// TIA Portal project "SludeProcess_Near_Final" (V16)

(* hardware
DEVICE "S71500/ET200MP station_1"  S7-1500 station
   slot 0: "Rail_0"  Rack  6ES7 590-1***0-0AA0
   slot 1: "PLC_1"  CPU 1511-1 PN  6ES7 511-1AK01-0AB0  V2.8
      slot 3: "CPU display_1"  6ES7591-1AA00-0AA0
      slot 32768: "PROFINET interface_1"  X1
         slot 32769: "Port_1"  X1 P1
         slot 32770: "Port_2"  X1 P2
      slot 34817: "Virtual CP interface port_1"  Virtual CP interface port  Virtual CP interface port
   slot 2: "DI 16x24VDC BA_1"  DI 16x24VDC BA  6ES7 521-1BH10-0AA0  V1.1
   slot 3: "DQ 16x24VDC/0.5A BA_1"  DQ 16x24VDC/0.5A BA  6ES7 522-1BH10-0AA0  V1.1
   slot 4: "AI 8xU/I/RTD/TC ST_1"  AI 8xU/I/RTD/TC ST  6ES7 531-7KF00-0AB0  V2.2
   slot 5: "AQ 2xU/I ST_1"  AQ 2xU/I ST  6ES7 532-5NB00-0AB0  V1.0
   slot 6: "DI 16x24VDC BA_2"  DI 16x24VDC BA  6ES7 521-1BH10-0AA0  V1.1
DEVICE "HMI_1"  KTP700 Basic PN
   slot 0: "HMI_1"  KTP700 Basic PN  6AV2 123-2GB03-0AX0  16.0.0.0
   slot 1: "HMI_RT_1"  KTP700 Basic PN  6AV2 123-2GB03-0AX0  16.0.0.0
   slot 5: "HMI_1.IE_CP_1"  PROFINET Interface  16.0.0.0
      slot 1: "PROFINET Interface_1"  PROFINET Interface
         slot 1: "Port_1"  Port
*)

// ===== PLC "PLC_1"  CPU 1511-1 PN =====

VAR_GLOBAL   // PLC tag table "Default tag table"
   "M001start" AT %M2.0 : Bool;
   "M001stop" AT %M12.1 : Bool;
   "FT-516_l/s" AT %MD12 : Real;
   "FT-516_status" AT %MW16 : Word;
   "FIC-516_setpoint" AT %MD18 : Real;
   "FIC-516_reset" AT %M2.1 : Bool;
   "M003_status" AT %MW20 : Word;
   "Test_open_valves" AT %M2.2 : Bool;
   "Test_M003_start" AT %M2.3 : Bool;
   "LT-515_liters" AT %MD22 : Real;
   "LT-515_status" AT %MW24 : Word;
   "M002_startbutton" AT %M2.4 : Bool;
   "M002_stopbutton" AT %M2.5 : Bool;
   "M002start" AT %M2.6 : Bool;
   "M002stop" AT %M2.7 : Bool;
   "WT-512_kg" AT %MD26 : Real;
   "TT-517_C" AT %MD28 : Real;
   "TT-518_C" AT %MD32 : Real;
   "WT-512_status" AT %MW36 : Word;
   "TT-517_status" AT %MW38 : Word;
   "TT-518_status" AT %MW40 : Word;
   "StartButton" AT %M3.0 : Bool;
   "StopButton" AT %M3.1 : Bool;
   "mixing" AT %M3.2 : Bool;
   "LSA513_HighLevel" AT %M3.3 : Bool;
   "HS519_FlowSwitch" AT %M3.4 : Bool;
   "HS514_MixReady" AT %M3.5 : Bool;
   "HS510_Valve" AT %M3.6 : Bool;
   "HS511_Valve" AT %M3.7 : Bool;
   "HS514_Valve" AT %M4.0 : Bool;
   "HS519_Valve" AT %M4.1 : Bool;
   "HS521_Alarm" AT %M4.2 : Bool;
   "M001_pMotor" AT %M4.3 : Bool;
   "M002_mix" AT %M4.4 : Bool;
   "M003_transferPump" AT %M4.5 : Bool;
   "FrequencyCommand" AT %MD42 : Real;
   "CurrentStep" AT %MW46 : Int;
   "Alarm" AT %M4.6 : Bool;
   "Step" AT %MW48 : Int;
   "NextStep" AT %MW50 : Int;
   "ResetButton" AT %M5.0 : Bool;
   "EmergencyButton" AT %M5.1 : Bool;
   "prevStart" AT %M5.2 : Bool;
   "prevStop" AT %M5.3 : Bool;
END_VAR

VAR_GLOBAL   // PLC tag table "SIMIT interface"
   "ZSO-510" AT %I0.0 : Bool;
   "ZSC-510" AT %I0.1 : Bool;
   "ZSO-511" AT %I0.2 : Bool;
   "ZSC-511" AT %I0.3 : Bool;
   "ZSO-514" AT %I0.4 : Bool;
   "ZSC-514" AT %I0.5 : Bool;
   "ZSO-519" AT %I0.6 : Bool;
   "ZSC-519" AT %I0.7 : Bool;
   "ZSO-521" AT %I1.0 : Bool;
   "ZSC-521" AT %I1.1 : Bool;
   "M001.R" AT %I1.2 : Bool;
   "M002.R" AT %I1.3 : Bool;
   "LS-513" AT %I1.4 : Bool;
   "GSV-510" AT %Q0.0 : Bool;
   "GSV-511" AT %Q0.1 : Bool;
   "GSV-514" AT %Q0.2 : Bool;
   "GSV-519" AT %Q0.3 : Bool;
   "GSV-521" AT %Q0.4 : Bool;
   "M001.ST" AT %Q0.5 : Bool;
   "M002.ST" AT %Q0.6 : Bool;
   "WT-512" AT %IW2 : Int;
   "LT-515" AT %IW4 : Int;
   "FT-516" AT %IW6 : Int;
   "TT-517" AT %IW8 : Int;
   "TT-518" AT %IW10 : Int;
   "M003.SP" AT %QW2 : Int;
   "M001.F" AT %I1.5 : Bool;
   "M002.F" AT %I1.6 : Bool;
   "M003.R" AT %I1.7 : Bool;
   "M003.F" AT %I18.0 : Bool;
   "M003.ST" AT %Q0.7 : Bool;
   "M001.TK" AT %I18.1 : Bool;
   "M002.TK" AT %I18.2 : Bool;
   "M003.TK" AT %I18.3 : Bool;
END_VAR

DATA_BLOCK "fb_ProcessSequence1_DB"   // DB2
{ S7_Optimized_Access := 'TRUE' }
VERSION : 0.1
// stored: InstanceOfName fb_ProcessSequence1
"fb_ProcessSequence1"
BEGIN
END_DATA_BLOCK

DATA_BLOCK "FIC516_DB"   // DB3
{ S7_Optimized_Access := 'TRUE' }
VERSION : 0.1
// stored: InstanceOfName FIC516
"FIC516"
BEGIN
END_DATA_BLOCK

DATA_BLOCK "AI_handeling_DB"   // DB14
{ S7_Optimized_Access := 'TRUE' }
VERSION : 0.1
// stored: InstanceOfName AI_handeling
"AI_handeling"
BEGIN
END_DATA_BLOCK

// folder: System blocks/Program resources

DATA_BLOCK "tMix"   // DB4
{ S7_Optimized_Access := 'TRUE' }
AUTHOR : Simatic
FAMILY : IEC
NAME : IEC_TMR
VERSION : 1.0
// stored: InstanceOfName IEC_TIMER
"IEC_TIMER"
BEGIN
END_DATA_BLOCK

// folder: (top level)

FUNCTION_BLOCK "FIC516"   // FB1, FBD
{ S7_Optimized_Access := 'TRUE' }
VERSION : 0.1
BEGIN

REGION Network 1
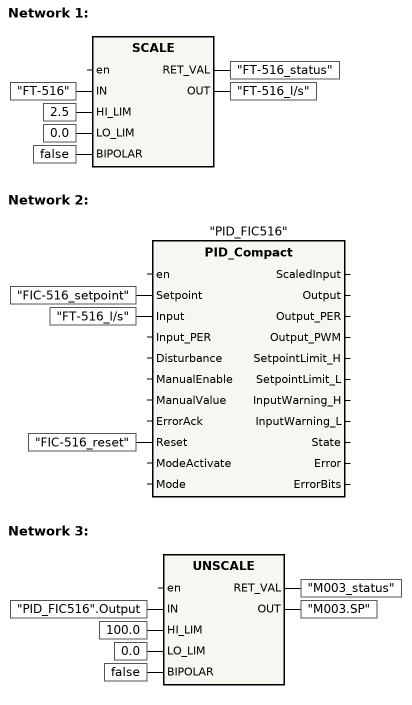
   "FT-516_status" := SCALE(IN := "FT-516", HI_LIM := 2.5, LO_LIM := 0.0, BIPOLAR := false, OUT => "FT-516_l/s");
END_REGION

REGION Network 2
   "PID_FIC516"(Setpoint := "FIC-516_setpoint", Input := "FT-516_l/s", Reset := "FIC-516_reset");   // PID_Compact
END_REGION

REGION Network 3
   "M003_status" := UNSCALE(IN := "PID_FIC516".Output,
                           HI_LIM := 100.0,
                           LO_LIM := 0.0,
                           BIPOLAR := false,
                           OUT => "M003.SP");
END_REGION
END_FUNCTION_BLOCK

FUNCTION_BLOCK "AI_handeling"   // FB4, FBD
{ S7_Optimized_Access := 'TRUE' }
VERSION : 0.1
BEGIN

REGION Network 1
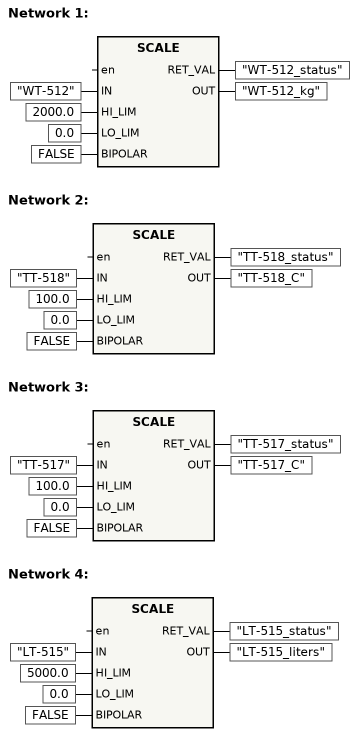
   "WT-512_status" := SCALE(IN := "WT-512",
                           HI_LIM := 2000.0,
                           LO_LIM := 0.0,
                           BIPOLAR := FALSE,
                           OUT => "WT-512_kg");
END_REGION

REGION Network 2
   "TT-518_status" := SCALE(IN := "TT-518", HI_LIM := 100.0, LO_LIM := 0.0, BIPOLAR := FALSE, OUT => "TT-518_C");
END_REGION

REGION Network 3
   "TT-517_status" := SCALE(IN := "TT-517", HI_LIM := 100.0, LO_LIM := 0.0, BIPOLAR := FALSE, OUT => "TT-517_C");
END_REGION

REGION Network 4
   "LT-515_status" := SCALE(IN := "LT-515",
                           HI_LIM := 5000.0,
                           LO_LIM := 0.0,
                           BIPOLAR := FALSE,
                           OUT => "LT-515_liters");
END_REGION
END_FUNCTION_BLOCK

FUNCTION_BLOCK "fb_ProcessSequence1"   // FB5, SCL
{ S7_Optimized_Access := 'TRUE' }
VERSION : 0.1
   VAR_INPUT
      StartButton : Bool := false;
      StopButton : Bool;
      RestartButton : Bool;
      ResetButton : Bool;
      EmergencyButton : Bool;
      "WT-512_kg" : Real;
      LT_515_liters : Real;
      FIC_516_setpoint : Real;
      TT_517_C : Real;
      TT_518_C : Real;
      LSA513_HighLevel : Bool;
      HS519_FlowSwitch : Bool;
      HS514_MixReady : Real;
      M001_SafetySwitch : Bool;
      M002_SafetySwitch : Bool;
      M003_SafetySwitch : Bool;
      Mode_Manual : Bool;
   END_VAR
   VAR_OUTPUT
      HS514_Valve : Bool;
      HS510_Valve : Bool;
      HS511_Valve : Bool;
      HS519_Valve : Bool;
      HS521_Valve : Bool;
      M001_pMotor : Bool;
      M002_mix : Bool;
      M003_TransferPump : Bool;
      FrequencyCommand : Real;
   END_VAR
   VAR
      Filling : Bool;
      WeightSetpoint : Real := 800.0;
      prevStart : Bool;
      AlarmActive : Bool;
      DosingNaOH : Bool;
      FeedingPowder : Bool;
      prevStop : Bool;
      Mixing : Bool;
      Transferring : Bool;
      StepMem : Bool;
      tMixTimer : Time;
      tFlowTimer : Time;
      "Step" : Int;
      Mode_Auto : Bool := true;
      HS519_manualValve : Bool;
      CircActive : Bool := false;
      MAN_HS510 : Bool;
      MAN_HS511 : Bool;
      MAN_HS514 : Bool;
      MAN_M001 : Bool;
      MAN_M002 : Bool;
      MAN_M003 : Bool;
      paused : Bool;
      M002_Fault_1 : Bool;
      restartLatch : Bool;
      TT_517_alarm : Bool;
      TT_518_alarm : Bool;
      LSA_513 : Bool := true;
      M001_Fault : Bool;
      M002_Fault : Bool;
      M003_Fault : Bool;
      CurrentStep : Int;
      Alarm : Bool;
      AlarmCause : String;
      M001_Safety : Bool;
      M002_Safety : Bool;
      M003_Safety : Bool;
      cMixTime : Time := T#20s;
      cOpenValveTime : Time := T#1000ms;
      cFlowCtrlTime : Time := T#50ms;
      running : Bool;
   END_VAR
   VAR CONSTANT
      cWeightWater : Real := 800.0;
      cWeightNaOH : Real := 1500.0;
      cWeightPowder : Real := 1000.0;
      cMaxWeight : Real := 2500.0;
      cFlowMin : Real := 0.5;
      cFlowMax : Real := 2.5;
      cTempEmergency : Real := 150.0;
      cTransferTrip : Real := 40.0;
      cFrequencyStep : Real := 1.0;
      cFrequenceMax : Real := 100.0;
      cFrequencyMin : Real;
   END_VAR
BEGIN
   // ---------- Immediate Emergency & Interlocks ----------
   IF #EmergencyButton OR (#TT_517_C >= #cTempEmergency) OR (#"WT-512_kg" >= #cMaxWeight) THEN
       #Alarm := TRUE;
       #AlarmCause := 'Emergency Stop or Max Temp/Weight Exceeded';
       #HS510_Valve := FALSE;
       #HS511_Valve := FALSE;
       #HS514_Valve := FALSE;
       #HS519_Valve := FALSE;
       #HS521_Valve := FALSE;
       #M001_pMotor := FALSE;
       #M002_mix := FALSE;
       #M003_TransferPump := FALSE;
       #FrequencyCommand := 0.0;
       #Step := 99;
       #paused := FALSE;
       RETURN;
   END_IF;

   // ---------- Default Outputs & HMI Indicators Initialization ----------
   // Hardware Outputs
   #HS510_Valve := FALSE;
   #HS511_Valve := FALSE;
   #HS514_Valve := FALSE;
   #HS519_Valve := FALSE;
   #HS521_Valve := FALSE;
   #M001_pMotor := FALSE;
   #M002_mix := FALSE;
   #M003_TransferPump := FALSE;
   #FrequencyCommand := 0.0;

   // HMI Status Indicators (Reset every scan, forced ON during active steps)
   #Filling := FALSE;
   #FeedingPowder := FALSE;
   #DosingNaOH := FALSE;
   #Mixing := FALSE;
   #Transferring := FALSE;
   #running := FALSE;

   // Automatic detection of motor faults & Alarms
   IF #TT_517_C >= #cTempEmergency THEN
       #TT_517_alarm := TRUE;
   END_IF;
   IF #TT_517_alarm THEN
       #M002_Fault := TRUE;
       #M002_Safety := FALSE;
       #Alarm := TRUE;
       #AlarmCause := 'TI-517 overtemp -> M002 fault';
   END_IF;

   IF #TT_518_C >= #cTempEmergency THEN
       #TT_518_alarm := TRUE;
   END_IF;
   IF #TT_518_alarm THEN
       #M003_Fault := TRUE;
       #M003_Safety := FALSE;
       #Alarm := TRUE;
       #AlarmCause := 'TI-518 overtemp -> M003 fault';
   END_IF;

   // LSA 513 Powder Hopper Low Level Warning
   IF NOT #LSA513_HighLevel AND (#AlarmCause = '') THEN
       #AlarmCause := 'LSA_513 Powder Hopper Low Level Warning';
   END_IF;

   // Reset alarm 
   IF #ResetButton THEN
       #Alarm := FALSE;
       #M001_Fault := FALSE;
       #M002_Fault := FALSE;
       #M003_Fault := FALSE;
       #TT_517_alarm := FALSE;
       #TT_518_alarm := FALSE;
       #AlarmCause := '';
   END_IF;

   // Restart (Only functions AFTER alarms are cleared)
   IF #RestartButton AND NOT #EmergencyButton AND NOT #Alarm THEN
       IF #M001_Safety AND #M002_Safety AND #M003_Safety AND NOT #M001_Fault AND NOT #M002_Fault AND NOT #M003_Fault THEN
           #Step := 0;
           #FrequencyCommand := 0.0;
           #paused := FALSE;
       END_IF;
   END_IF;

   // Hardware Safety Switch Mapping (TRUE = Healthy Motor)
   #M001_Safety := #M001_SafetySwitch;
   #M002_Safety := #M002_SafetySwitch;
   #M003_Safety := #M003_SafetySwitch;

   // Delivery Request mapping
   IF #HS519_FlowSwitch THEN
       #HS519_manualValve := TRUE;
   ELSE
       #HS519_manualValve := FALSE;
   END_IF;

   // ---------- Manual mode ----------
   IF #Mode_Manual THEN
       #running := TRUE;
       #Mode_Auto := FALSE;

       IF #MAN_HS510 AND #M001_Safety AND #M002_Safety THEN
           #HS510_Valve := TRUE;
           #Filling := TRUE;
       END_IF;
       IF #MAN_HS511 AND #M002_Safety THEN
           #HS511_Valve := TRUE;
           #DosingNaOH := TRUE;
       END_IF;
       IF #MAN_HS514 THEN
           #HS514_Valve := TRUE;
           #Transferring := TRUE;
       END_IF;

       IF #MAN_M001 AND NOT #M001_Fault AND #M001_Safety THEN
           #M001_pMotor := TRUE;
           #FeedingPowder := TRUE;
       END_IF;

       IF #MAN_M002 AND NOT #M002_Fault AND #M002_Safety THEN
           #M002_mix := TRUE;
           #Mixing := TRUE;
       END_IF;

       IF #MAN_M003 AND NOT #M003_Fault AND #M003_Safety THEN
           #M003_TransferPump := TRUE;
       END_IF;

       GOTO Global_Interlocks;
   END_IF;


   // ---------- Auto Sequence Controls ----------
   IF #StopButton AND (NOT #prevStop) THEN
       #paused := NOT #paused; // rising edge toggle
   END_IF;
   IF #StartButton THEN
       #paused := FALSE;
   END_IF;
   #prevStop := #StopButton;

   IF #paused THEN
       #AlarmCause := 'Process PAUSED';
       GOTO Global_Interlocks;
   ELSE
       IF #AlarmCause = 'Process PAUSED' THEN
           #AlarmCause := '';
       END_IF;
   END_IF;


   // ==============================================================================
   // INDEPENDENT STORAGE TANK BACKGROUND CIRCULATION (Runs constantly in Auto Mode)
   // ==============================================================================
   IF #Mode_Auto AND (#Step <> 99) THEN
       IF #LT_515_liters > 500.0 THEN
           IF #M003_Safety AND NOT #M003_Fault THEN
               #M003_TransferPump := TRUE;
               #running := TRUE;

               IF #HS519_manualValve THEN
                   // Delivery Mode Active
                   #HS519_Valve := TRUE;
                   #HS521_Valve := FALSE;
                   #CircActive := FALSE;

                   // Flow Control logic
                   IF #FIC_516_setpoint > #cFlowMin AND #FIC_516_setpoint < #cFlowMax THEN
                       IF #FrequencyCommand < #FIC_516_setpoint THEN
                           #FrequencyCommand := MIN(IN1 := #FrequencyCommand + #cFrequencyStep, IN2 := #cFrequenceMax);
                       ELSIF #FrequencyCommand > #FIC_516_setpoint THEN
                           #FrequencyCommand := MAX(IN1 := #FrequencyCommand - #cFrequencyStep, IN2 := #cFrequencyMin);
                       END_IF;
                   END_IF;
               ELSE
                   // Default Recirculation Mode Active
                   #HS519_Valve := FALSE;
                   #HS521_Valve := TRUE;
                   #CircActive := TRUE;
               END_IF;
           ELSE
               #M003_TransferPump := FALSE;
               #CircActive := FALSE;
               #Alarm := TRUE;
               #AlarmCause := 'M003 unsafe for delivery/recirculation';
               #Step := 99;
           END_IF;
       END_IF;
   END_IF;
   // ==============================================================================


   // ---------- State Machine (Mix Tank Batching Sequence) ----------
   CASE #Step OF

       0: // Standby
           #Mode_Auto := TRUE;
           IF #StartButton THEN
               #Step := 2;
           END_IF;

       2: // Start Check
           #Mode_Auto := TRUE;
           IF #Mode_Auto THEN
               #Step := 3;
               "tMix".TON(IN := FALSE,
                          PT := #cMixTime); // Hard reset the timer so it is fresh for the new batch
           ELSE
               IF #StartButton THEN
                   #running := TRUE;
               END_IF;
           END_IF;

       3: // Water Dosing (HS 510)
           IF #M001_Safety AND NOT #M002_Fault THEN
               #HS510_Valve := TRUE;
               #running := TRUE;
               #Filling := TRUE;
           ELSE
               #Alarm := TRUE;
               #AlarmCause := 'Equipment unsafe for water fill';
               #Step := 99;
           END_IF;

           IF #"WT-512_kg" >= #cWeightWater THEN
               #Step := 4;
           END_IF;

       4: // Powder Dosing & Mixing (M001 & M002)
           IF #M001_Safety AND #M002_Safety AND NOT #M001_Fault AND NOT #M002_Fault THEN
               #M001_pMotor := TRUE;
               #M002_mix := TRUE;
               #FeedingPowder := TRUE;
               #Mixing := TRUE;
               #running := TRUE;
           ELSE
               #Alarm := TRUE;
               #AlarmCause := 'M001/M002 safety fault prevented powder feed';
               #Step := 99;
           END_IF;

           IF #"WT-512_kg" >= #cWeightPowder THEN
               #Step := 5;
           END_IF;

       5: // Sodium Hydroxide Dosing (HS 511 & M002)
           IF #M002_Safety AND NOT #M002_Fault THEN
               #HS511_Valve := TRUE;
               #M002_mix := TRUE;
               #DosingNaOH := TRUE;
               #Mixing := TRUE;
               #running := TRUE;
           ELSE
               #Alarm := TRUE;
               #AlarmCause := 'M002 unsafe during NaOH dosing';
               #Step := 99;
           END_IF;

           IF #"WT-512_kg" >= #cWeightNaOH THEN
               #Step := 6;
           END_IF;

       6: // Final Mixing Time (Waits for proper mix before transfer)
           IF #M002_Safety AND NOT #M002_Fault THEN
               #M002_mix := TRUE;
               #Mixing := TRUE;
               #running := TRUE;

               // Run the TON Timer
               "tMix".TON(IN := TRUE,
                          PT := #cMixTime,
                          ET => #tMixTimer);
           ELSE
               #Alarm := TRUE;
               #AlarmCause := 'M002 unsafe for final mixing';
               #Step := 99;
           END_IF;

           // Once the timer hits the PT value (e.g., 5s), Q goes TRUE
           IF "tMix".Q THEN
               "tMix".TON(IN := FALSE,
                          PT := #cMixTime); // Reset the timer before moving on
               #Step := 7;
           END_IF;

       7: // Transfer to Storage Tank (HS 514)
           IF #LT_515_liters < 4950.0 THEN
               #HS514_Valve := TRUE;
               #running := TRUE;
               #Transferring := TRUE;
           END_IF;

           // Sequence finishes when Mix Tank is empty. Goes straight back to Standby!
           IF (#"WT-512_kg" <= 10.0) OR (#LT_515_liters >= 4950.0) THEN
               #Step := 0;
           END_IF;

       99: // Fault State
           #running := FALSE;
           #CircActive := FALSE;

           // 1. Operator MUST press Reset first to clear the alarm
           IF #ResetButton THEN
               IF #M001_SafetySwitch AND #M002_SafetySwitch AND #M003_SafetySwitch AND NOT #M001_Fault AND NOT #M002_Fault AND NOT #M003_Fault THEN
                   #Alarm := FALSE; // Fault cleared successfully
                   #AlarmCause := '';
               ELSE
                   #Alarm := TRUE;
                   #AlarmCause := 'Cannot clear emergency - check faults/safety';
               END_IF;
           END_IF;

           // 2. ONLY after Reset clears the alarm, wait for Start or Restart command
           IF NOT #Alarm THEN
               IF #StartButton THEN
                   #Step := 2; // Press START to resume the batch from where it failed
               ELSIF #RestartButton THEN
                   #Step := 0; // Press RESTART to abort batch and return to Standby
               END_IF;
           END_IF;

       ELSE
           #Step := 0;
   END_CASE;

   // ---------- Global Interlocks (Applies to both Auto & Manual) ----------
   Global_Interlocks:

   // 1. Storage Tank Overflow Protection
   IF #LT_515_liters >= 4950.0 THEN
       #HS514_Valve := FALSE;
   END_IF;

   // 2. Storage Tank Low Level Pump Protection
   IF #LT_515_liters <= 500.0 THEN
       #M003_TransferPump := FALSE;
       #HS521_Valve := FALSE;
       #HS519_Valve := FALSE;
   END_IF;

   // 3. Flow Diverter Interlock: Cannot be open at the same time
   IF #HS519_Valve AND #HS521_Valve THEN
       #HS521_Valve := FALSE;
   END_IF;

   #CurrentStep := #Step;
END_FUNCTION_BLOCK

ORGANIZATION_BLOCK "Main"   // OB1, FBD, ProgramCycle
TITLE = "Main Program Sweep (Cycle)"
{ S7_Optimized_Access := 'TRUE' }
VERSION : 0.1
   VAR_INPUT
      Initial_Call : Bool;   // Initial call of this OB
      Remanence : Bool;   // =True, if remanent data are available
   END_VAR
BEGIN

REGION Network 1
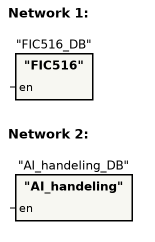
   "FIC516_DB"();   // "FIC516"
END_REGION

REGION Network 2
   "AI_handeling_DB"();   // "AI_handeling"
END_REGION

REGION Network 3
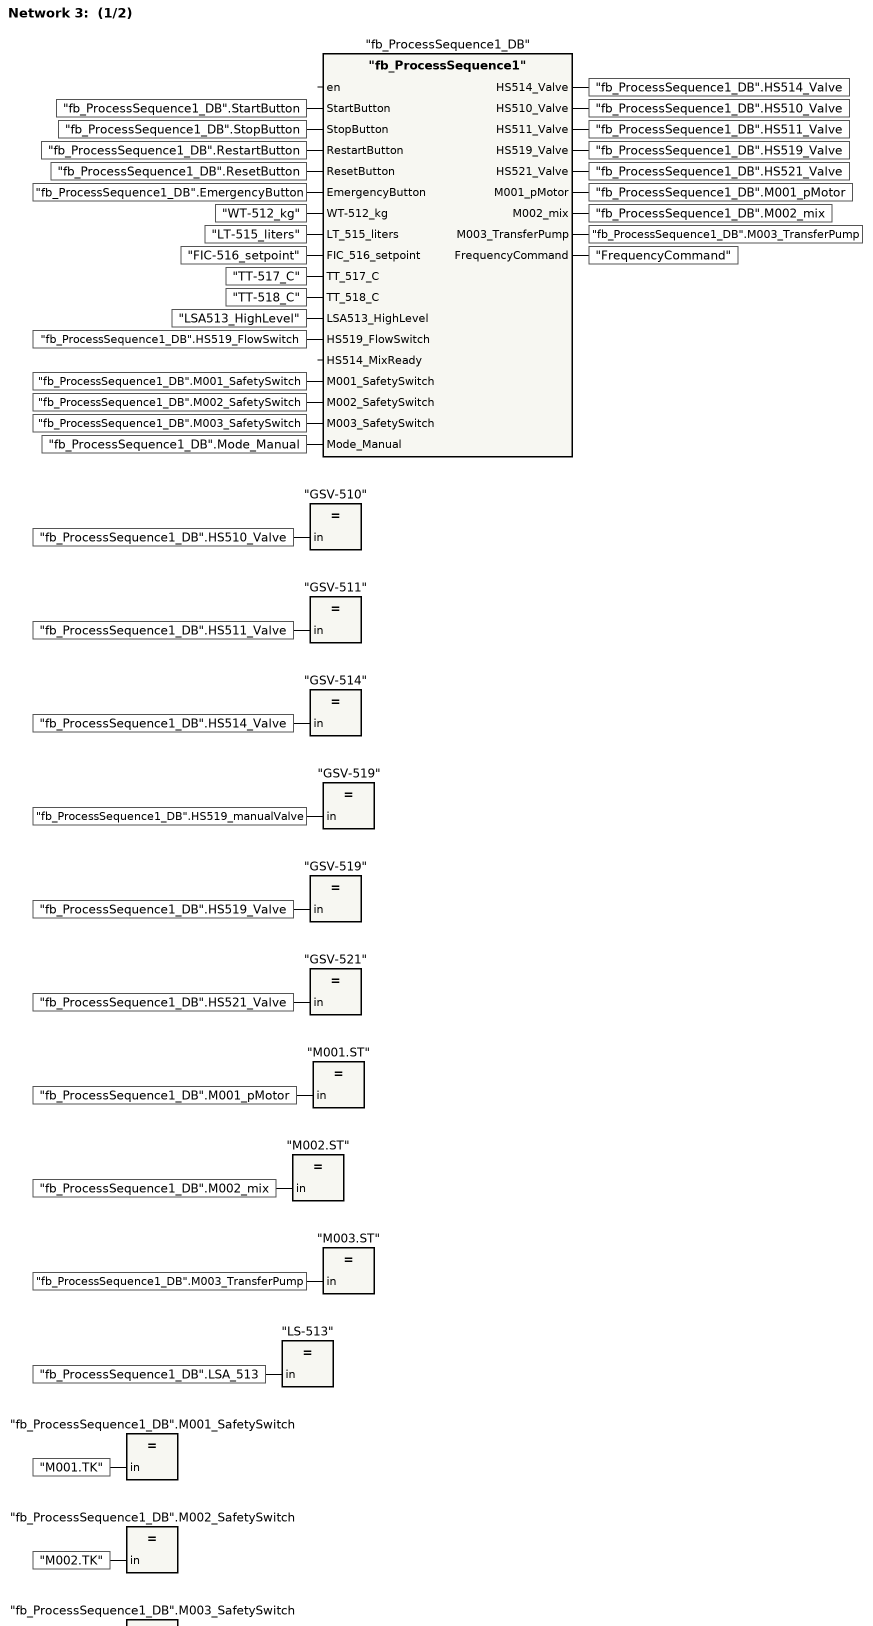
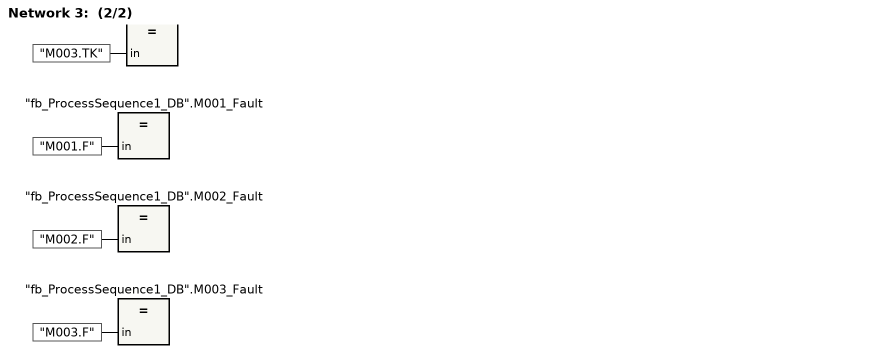
   "fb_ProcessSequence1_DB"(StartButton := "fb_ProcessSequence1_DB".StartButton,   // "fb_ProcessSequence1"
                           StopButton := "fb_ProcessSequence1_DB".StopButton,
                           RestartButton := "fb_ProcessSequence1_DB".RestartButton,
                           ResetButton := "fb_ProcessSequence1_DB".ResetButton,
                           EmergencyButton := "fb_ProcessSequence1_DB".EmergencyButton,
                           "WT-512_kg" := "WT-512_kg",
                           LT_515_liters := "LT-515_liters",
                           FIC_516_setpoint := "FIC-516_setpoint",
                           TT_517_C := "TT-517_C",
                           TT_518_C := "TT-518_C",
                           LSA513_HighLevel := "LSA513_HighLevel",
                           HS519_FlowSwitch := "fb_ProcessSequence1_DB".HS519_FlowSwitch,
                           M001_SafetySwitch := "fb_ProcessSequence1_DB".M001_SafetySwitch,
                           M002_SafetySwitch := "fb_ProcessSequence1_DB".M002_SafetySwitch,
                           M003_SafetySwitch := "fb_ProcessSequence1_DB".M003_SafetySwitch,
                           Mode_Manual := "fb_ProcessSequence1_DB".Mode_Manual,
                           HS514_Valve => "fb_ProcessSequence1_DB".HS514_Valve,
                           HS510_Valve => "fb_ProcessSequence1_DB".HS510_Valve,
                           HS511_Valve => "fb_ProcessSequence1_DB".HS511_Valve,
                           HS519_Valve => "fb_ProcessSequence1_DB".HS519_Valve,
                           HS521_Valve => "fb_ProcessSequence1_DB".HS521_Valve,
                           M001_pMotor => "fb_ProcessSequence1_DB".M001_pMotor,
                           M002_mix => "fb_ProcessSequence1_DB".M002_mix,
                           M003_TransferPump => "fb_ProcessSequence1_DB".M003_TransferPump,
                           FrequencyCommand => "FrequencyCommand");
   "GSV-510" := "fb_ProcessSequence1_DB".HS510_Valve;
   "GSV-511" := "fb_ProcessSequence1_DB".HS511_Valve;
   "GSV-514" := "fb_ProcessSequence1_DB".HS514_Valve;
   "GSV-519" := "fb_ProcessSequence1_DB".HS519_manualValve;
   "GSV-519" := "fb_ProcessSequence1_DB".HS519_Valve;
   "GSV-521" := "fb_ProcessSequence1_DB".HS521_Valve;
   "M001.ST" := "fb_ProcessSequence1_DB".M001_pMotor;
   "M002.ST" := "fb_ProcessSequence1_DB".M002_mix;
   "M003.ST" := "fb_ProcessSequence1_DB".M003_TransferPump;
   "LS-513" := "fb_ProcessSequence1_DB".LSA_513;
   "fb_ProcessSequence1_DB".M001_SafetySwitch := "M001.TK";
   "fb_ProcessSequence1_DB".M002_SafetySwitch := "M002.TK";
   "fb_ProcessSequence1_DB".M003_SafetySwitch := "M003.TK";
   "fb_ProcessSequence1_DB".M001_Fault := "M001.F";
   "fb_ProcessSequence1_DB".M002_Fault := "M002.F";
   "fb_ProcessSequence1_DB".M003_Fault := "M003.F";
END_REGION
END_ORGANIZATION_BLOCK

ORGANIZATION_BLOCK "Startup"   // OB100, SCL, Startup
TITLE = "Complete Restart"
{ S7_Optimized_Access := 'TRUE' }
VERSION : 0.1
   VAR_INPUT
      LostRetentive : Bool;   // True if retentive data are lost
      LostRTC : Bool;   // True if date and time are lost
   END_VAR
BEGIN
   (* dEFAULT FLOW SETPOINT VALUE*)
   "Step" := 0;

   "FIC-516_setpoint" := 0.5;
END_ORGANIZATION_BLOCK

(* ===== HMI "HMI_RT_1" =====
system functions are stored by id; their names below are inferred from use
connection "HMI_Connection_1": ETHERNET, SMART_S7_1500_OMS

HMI tags "Default tag table"
   "fb_processSequence_DB_Alarm" : Bool = PLC fb_ProcessSequence1_DB.Alarm AT %M4.6, 1 s
   "fb_processSequence_DB_AlarmCause" : String[254] = PLC fb_ProcessSequence1_DB.AlarmCause AT %M4.6, 1 s
   "fb_processSequence_DB_EmergencyButton" : Bool = PLC fb_ProcessSequence1_DB.EmergencyButton AT %M5.1, 1 s
   "fb_processSequence_DB_FIC_516_setpoint" : Real = PLC fb_ProcessSequence1_DB.FIC_516_setpoint AT %MD18, 1 s
   "fb_processSequence_DB_HS510_Valve" : Bool = PLC fb_ProcessSequence1_DB.HS510_Valve AT %DB1.DBX0.0, 1 s
   "fb_processSequence_DB_HS511_Valve" : Bool = PLC fb_ProcessSequence1_DB.HS511_Valve AT %Q0.1, 1 s
   "fb_processSequence_DB_HS514_Valve" : Bool = PLC fb_ProcessSequence1_DB.HS514_Valve AT %Q0.2, 1 s
   "fb_processSequence_DB_HS519_FlowSwitch" : Bool = PLC fb_ProcessSequence1_DB.HS519_FlowSwitch AT %M3.4, 1 s
   "fb_processSequence_DB_HS519_manualValve" : Bool = PLC fb_ProcessSequence1_DB.HS519_manualValve AT %M4.1, 1 s
   "fb_processSequence_DB_LT-515_liters" : Real = PLC fb_ProcessSequence1_DB.LT_515_liters AT %MD22, 1 s
   "fb_processSequence_DB_M001_pMotor" : Bool = PLC fb_ProcessSequence1_DB.M001_pMotor AT %M4.3, 1 s
   "fb_processSequence_DB_M002_mix" : Bool = PLC fb_ProcessSequence1_DB.M002_mix AT %M4.4, 1 s
   "fb_processSequence_DB_MAN_HS510" : Bool = PLC fb_ProcessSequence1_DB.MAN_HS510 AT %M3.6, 1 s
   "fb_processSequence_DB_MAN_HS511" : Bool = PLC fb_ProcessSequence1_DB.MAN_HS511 AT %M3.7, 1 s
   "fb_processSequence_DB_MAN_HS514" : Bool = PLC fb_ProcessSequence1_DB.MAN_HS514 AT %M4.0, 1 s
   "fb_processSequence_DB_MAN_M001" : Bool = PLC fb_ProcessSequence1_DB.MAN_M001 AT %DB1.DBX0.0, 1 s
   "fb_processSequence_DB_MAN_M002" : Bool = PLC fb_ProcessSequence1_DB.MAN_M002 AT %DB1.DBX0.0, 1 s
   "fb_processSequence_DB_MAN_M003" : Bool = PLC fb_ProcessSequence1_DB.MAN_M003 AT %DB1.DBX0.0, 1 s
   "fb_processSequence_DB_Mixing" : Bool = PLC fb_ProcessSequence1_DB.Mixing AT %DB1.DBX0.0, 1 s
   "fb_processSequence_DB_Mode_Auto" : Bool = PLC fb_ProcessSequence1_DB.Mode_Auto AT %DB1.DBX0.0, 1 s
   "fb_processSequence_DB_Mode_Manual" : Bool = PLC fb_ProcessSequence1_DB.Mode_Manual AT %DB1.DBX0.0, 1 s
   "fb_processSequence_DB_ResetButton" : Bool = PLC fb_ProcessSequence1_DB.ResetButton AT %DB1.DBX0.0, 1 s
   "fb_processSequence_DB_RestartButton" : Bool = PLC fb_ProcessSequence1_DB.RestartButton AT %DB1.DBX0.0, 1 s
   "fb_processSequence_DB_running" : Bool = PLC fb_ProcessSequence1_DB.running AT %DB1.DBX0.0, 1 s
   "fb_processSequence_DB_StartButton" : Bool = PLC fb_ProcessSequence1_DB.StartButton AT %DB1.DBX0.0, 1 s
   "fb_processSequence_DB_StopButton" : Bool = PLC fb_ProcessSequence1_DB.StopButton AT %DB1.DBX0.0, 1 s
   "FIC-516_setpoint" : Real = PLC "FIC-516_setpoint" AT %MD18, 1 s
   "FT-516_l/s" : Real = PLC "FT-516_l/s" AT %MD12, 1 s
   "Tag_ScreenNumber" : UInt, internal

Template "Template_1" 800x480
   Button "Exit" at 714,429 size 71x50; TextOff 'Exit'; PictureOff "ExitRuntime_KTP700_Basic_PN_TR"; PictureOn "ExitRuntime_KTP700_Basic_PN_TR"
      on Release: StopRuntime(0)
   Button "Template_Button" at 614,429 size 71x50; TextOff 'Text'
   Button "Template_Button_1" at 514,429 size 71x50; TextOff 'Text'
   Button "Template_Button_2" at 414,429 size 71x50; TextOff 'Text'
   Button "Template_Button_3" at 314,429 size 71x50; TextOff 'Text'
   Button "Template_Button_4" at 214,429 size 71x50; TextOff 'Text'
   Button "Template_Button_5" at 114,429 size 71x50; TextOff 'Text'
      on Release: function_ef3f5d25("Alarm window_Unacknowledged", -1)
   Button "Start screen" at 14,422 size 71x50; TextOff 'Start screen'; PictureOff "NavigateHome_KTP700_Basic_PN_TR"; PictureOn "NavigateHome_KTP700_Basic_PN_TR"
      on Release: ActivateScreen("Root screen", 0)
   SymbolicIOField "Symbolic_IO_Field_Screen" at 93,9 size 600x33; TextOff '0'; TextOn '1'; TextList "TextList_ScreenNames"
      on Change: ActivateScreenByNumber("Tag_ScreenNumber", 0)
   DateTimeField "HmiScreenItemData" at 695,25 size 105x25
   DateTimeField "HmiScreenItemData_1" at 695,0 size 105x25
   GraphicView "Logo" at 0,0 size 91x51; Picture "Logo of HMI_1"

screen "Root screen" 800x480, template "Template_1"
   on GenerateScreen: SetTag("Tag_ScreenNumber", 1)
   IOField "I/O field_1" at 3,360 size 96x32; FormatPattern 9.99
      ProcessValue <- "FT-516_l/s"
   TextField "Text field_1" at 0,391 size 122x23; Text 'MEASURMENT'
   IOField "I/O field_2" at 3,280 size 96x32; FormatPattern 9.99
      ProcessValue <- "FIC-516_setpoint"
   TextField "Text field_2" at 5,315 size 89x23; Text 'SETPOINT'
   Circle "Circle_1" at 325,93 size 28x28
      Visibility <- "fb_processSequence_DB_StopButton"
   Switch "Switch_1" at 4,81 size 56x21; CaptionText 'Switch'; TextOff 'OFF'; TextOn 'ON'
      ProcessValue <- "fb_processSequence_DB_MAN_HS510"
   TextField "Text field_3" at 3,55 size 57x23; Text 'HS510'
   TextField "Text field_4" at 3,109 size 57x23; Text 'HS511'
   Switch "Switch_2" at 6,133 size 56x21; TextOn 'ON'; CaptionText 'Switch'; TextOff 'OFF'
      ProcessValue <- "fb_processSequence_DB_MAN_HS511"
   TextField "Text field_5" at 5,176 size 57x23; Text 'HS514'
   Switch "Switch_3" at 3,199 size 56x21; TextOn 'ON'; CaptionText 'Switch'; TextOff 'OFF'
      ProcessValue <- "fb_processSequence_DB_MAN_HS514"
   Circle "Circle_5" at 414,93 size 28x28
      Visibility <- "fb_processSequence_DB_RestartButton"
   Switch "Switch_6" at 79,80 size 56x21; TextOn 'ON'; CaptionText 'Switch'; TextOff 'OFF'
      ProcessValue <- "fb_processSequence_DB_MAN_M001"
   TextField "Text field_6" at 73,55 size 49x23; Text 'M002'
   TextField "Text field_7" at 161,57 size 49x23; Text 'M001'
   Switch "Switch_7" at 163,78 size 56x21; TextOn 'ON'; CaptionText 'Switch'; TextOff 'OFF'
      ProcessValue <- "fb_processSequence_DB_MAN_M001"
   Circle "Circle_6" at 506,93 size 28x28
      Visibility <- "fb_processSequence_DB_ResetButton"
   TextField "Text field_8" at 78,109 size 49x23; Text 'M003'
   Switch "Switch_8" at 78,133 size 56x21; TextOn 'ON'; CaptionText 'Switch'; TextOff 'OFF'
      ProcessValue <- "fb_processSequence_DB_MAN_M003"
   Circle "Circle_8" at 245,91 size 28x28
      Visibility <- "fb_processSequence_DB_StartButton"
   Switch "Switch_9" at 78,202 size 56x21; TextOn 'ON'; CaptionText 'Switch'; TextOff 'OFF'
      ProcessValue <- "fb_processSequence_DB_HS519_manualValve"
   TextField "Text field_11" at 78,174 size 57x23; Text 'HS519'
   TextField "Text field_9" at 252,384 size 115x23; Text 'Storage Tank'
   Circle "Circle_2" at 537,146 size 28x28
      Visibility <- "fb_processSequence_DB_Mode_Manual"
   Circle "Circle_3" at 537,202 size 28x28
      Visibility <- "fb_processSequence_DB_Mode_Auto"
   Circle "Circle_4" at 537,251 size 28x28
      Visibility <- "fb_processSequence_DB_Alarm"
   Circle "Circle_7" at 537,296 size 28x28
      Visibility <- "fb_processSequence_DB_running"
   Circle "Circle_9" at 607,90 size 28x28
      Visibility <- "fb_processSequence_DB_EmergencyButton"
   TextField "Text field_18" at 584,146 size 129x23; Text 'MANUAL MODE'
   TextField "Text field_19" at 574,202 size 100x23; Text 'AUTOMODE'
   TextField "Text field_20" at 583,254 size 58x23; Text 'FAULT'
   TextField "Text field_21" at 583,303 size 89x23; Text 'RUNNUNG'
   Circle "Circle_10" at 537,338 size 28x28
      Visibility <- "fb_processSequence_DB_Mixing"
   TextField "Text field_22" at 590,347 size 68x23; Text 'MIXING'
   Switch "Switch_4" at 449,148 size 56x21; TextOn 'ON'; CaptionText 'Switch'; TextOff 'OFF'
      ProcessValue <- "fb_processSequence_DB_Mode_Manual"
   Switch "Switch_5" at 274,198 size 56x21; TextOn 'ON'; CaptionText 'Switch'; TextOff 'OFF'
      ProcessValue <- "fb_processSequence_DB_HS519_FlowSwitch"
   TextField "Text field_23" at 445,166 size 68x23; Text 'ON/OFF'
   Bar "Bar_1" at 265,229 size 87x154; MinimumValue 0; MaximumValue 5000
      ProcessValue <- "fb_processSequence_DB_LT-515_liters"
   TextField "Text field_24" at 222,175 size 16x23; Text 'Text'
   Button "Button_1" at 229,65 size 74x25; TextOff 'START'
      on Press: SetBit("fb_processSequence_DB_StartButton")
      on Release: ResetBit("fb_processSequence_DB_StartButton")
   Button "Button_2" at 576,64 size 104x25; TextOff 'EMERGENCY'
      on Press: SetBit("fb_processSequence_DB_EmergencyButton")
      on Release: ResetBit("fb_processSequence_DB_EmergencyButton")
   Button "Button_3" at 484,63 size 74x25; TextOff 'RESET'
      on Press: SetBit("fb_processSequence_DB_ResetButton")
      on Release: ResetBit("fb_processSequence_DB_ResetButton")
   Button "Button_4" at 385,65 size 84x25; TextOff 'RESTART'
      on Press: SetBit("fb_processSequence_DB_RestartButton")
      on Release: ResetBit("fb_processSequence_DB_RestartButton")
   Button "Button_5" at 308,65 size 74x25; TextOff 'STOP'
      on Press: SetBit("fb_processSequence_DB_StopButton")
      on Release: ResetBit("fb_processSequence_DB_StopButton")
   TextField "Text field_10" at 248,174 size 107x23; Text 'Process flow'
*)